FUNCTION_BLOCK FB_CIP_Client EXTENDS FB_SFC_Cycle IMPLEMENTS ITF_FB_SFC_Cycle
VAR_INPUT
	//eElementID			: E_Element_List;
	
	valClient_Source		: E_Pis_Name;
	valClient_Return		: E_Pis_Name;
	valS_Marinade_Up		: E_Pis_Name;
	//valS_Marinade_Up_Drain	: E_Pis_Name;
	valS_Marinade_Low		: E_Pis_Name;
	valS_Color_Up			: E_Pis_Name;
	//valS_Color_Up_Drain		: E_Pis_Name;
	valS_Color_Low			: E_Pis_Name;
	//valTank_1				: E_Pis_Name;
	//valTank_2				: E_Pis_Name;
	//valTank_3				: E_Pis_Name;
	//valTank_4				: E_Pis_Name;
	//valS_Marinade_Low_Select	: E_Pis_Name;
	//valS_Color_Low_Select	: E_Pis_Name;
	valDrain				: E_Pis_Name;
	valLoop					: E_Pis_Name;//V1030
	valS_Future				: E_Pis_Name;
	
END_VAR
VAR_OUTPUT
END_VAR
VAR
	//refElement		: REFERENCE TO FB_Element;
	//refState_Long		: REFERENCE TO E_Element_State_Long;
	eReq				: E_CIP_Client_Selector;
	eProcess			: E_CIP_Client_Selector;
	eStatus				: E_CIP_Client_Selector;
	
	fbPis					: FB_Piston;
	stPis_Client_Source			: REFERENCE TO ST_Piston;
	stPis_Client_Return			: REFERENCE TO ST_Piston;
	stPis_S_Marinade_Up			: REFERENCE TO ST_Piston;
	//stPis_S_Marinade_Up_Drain	: REFERENCE TO ST_Piston;
	stPis_S_Marinade_Low		: REFERENCE TO ST_Piston;
	stPis_S_Color_Up			: REFERENCE TO ST_Piston;
	//stPis_S_Color_Up_Drain		: REFERENCE TO ST_Piston;
	stPis_S_Color_Low			: REFERENCE TO ST_Piston;
	//stPis_Tank_1				: REFERENCE TO ST_Piston;
	//stPis_Tank_2				: REFERENCE TO ST_Piston;
	//stPis_Tank_3				: REFERENCE TO ST_Piston;
	//stPis_Tank_4				: REFERENCE TO ST_Piston;
	//stPis_S_Marinade_Low_Select	: REFERENCE TO ST_Piston;
	//stPis_S_Color_Low_Select	: REFERENCE TO ST_Piston;
	stPis_Drain					: REFERENCE TO ST_Piston;	
	stPis_Loop					: REFERENCE TO ST_Piston;//V1030
	stPis_S_Future				: REFERENCE TO ST_Piston;

	tonDrainTime: TON;
	
	rt_Req_Reset: R_TRIG;

END_VAR
VAR_IN_OUT


END_VAR

act_GetReference();

act_Oper();
IF NOT Init.x THEN;
	act_Status();
END_IF

tonDrainTime(PT:=T#1M, IN:=eStatus=E_CIP_Client_Selector.eDrain);
IF tonDrainTime.Q 
AND eReq=E_CIP_Client_Selector.eNone
AND eProcess=E_CIP_Client_Selector.eNone
THEN;
	eReq:=E_CIP_Client_Selector.eClose;
END_IF

m_Request_Reset(memo:=rt_Req_Reset);//rt_Req_Reset: R_TRIG;

ACTION _aClose_active:
bStepDone:=FALSE;
IF TRUE 
AND eStatus=E_CIP_Client_Selector.eClose
THEN;
	bStepDone:=TRUE;
END_IF
END_ACTION

ACTION _aClose_entry:
fbPis.m_SetByRecipe(stPis:=stPis_Client_Source, 		req:=E_Piston_Recipe_State.Release);
fbPis.m_SetByRecipe(stPis:=stPis_Client_Return, 		req:=E_Piston_Recipe_State.Release);
fbPis.m_SetByRecipe(stPis:=stPis_S_Marinade_Up, 		req:=E_Piston_Recipe_State.Release);
fbPis.m_SetByRecipe(stPis:=stPis_S_Marinade_Low, 		req:=E_Piston_Recipe_State.Release);
fbPis.m_SetByRecipe(stPis:=stPis_S_Color_Up, 			req:=E_Piston_Recipe_State.Release);
fbPis.m_SetByRecipe(stPis:=stPis_S_Color_Low, 			req:=E_Piston_Recipe_State.Release);
fbPis.m_SetByRecipe(stPis:=stPis_Drain, 				req:=E_Piston_Recipe_State.Release);
fbPis.m_SetByRecipe(stPis:=stPis_Loop, 					req:=E_Piston_Recipe_State.Release);
fbPis.m_SetByRecipe(stPis:=stPis_S_Future, 				req:=E_Piston_Recipe_State.Release);
END_ACTION

ACTION _aColor_Low_active:
bStepDone:=FALSE;
IF TRUE 
AND eStatus=E_CIP_Client_Selector.eColor_Low
THEN;
	bStepDone:=TRUE;
END_IF
END_ACTION

ACTION _aColor_Low_entry:
fbPis.m_SetByRecipe(stPis:=stPis_Client_Source, 		req:=E_Piston_Recipe_State.Act);
fbPis.m_SetByRecipe(stPis:=stPis_Client_Return, 		req:=E_Piston_Recipe_State.Act);
fbPis.m_SetByRecipe(stPis:=stPis_S_Marinade_Up, 		req:=E_Piston_Recipe_State.Release);
fbPis.m_SetByRecipe(stPis:=stPis_S_Marinade_Low, 		req:=E_Piston_Recipe_State.Release);
fbPis.m_SetByRecipe(stPis:=stPis_S_Color_Up, 			req:=E_Piston_Recipe_State.Release);
fbPis.m_SetByRecipe(stPis:=stPis_S_Color_Low, 			req:=E_Piston_Recipe_State.Act);
fbPis.m_SetByRecipe(stPis:=stPis_Drain, 				req:=E_Piston_Recipe_State.Release);
fbPis.m_SetByRecipe(stPis:=stPis_Loop, 					req:=E_Piston_Recipe_State.Release);
fbPis.m_SetByRecipe(stPis:=stPis_S_Future, 				req:=E_Piston_Recipe_State.Release);
END_ACTION

ACTION _aColor_Up_active:
bStepDone:=FALSE;
IF TRUE 
AND eStatus=E_CIP_Client_Selector.eColor_Up
THEN;
	bStepDone:=TRUE;
END_IF
END_ACTION

ACTION _aColor_Up_entry:
fbPis.m_SetByRecipe(stPis:=stPis_Client_Source, 		req:=E_Piston_Recipe_State.Act);
fbPis.m_SetByRecipe(stPis:=stPis_Client_Return, 		req:=E_Piston_Recipe_State.Act);
fbPis.m_SetByRecipe(stPis:=stPis_S_Marinade_Up, 		req:=E_Piston_Recipe_State.Release);
fbPis.m_SetByRecipe(stPis:=stPis_S_Marinade_Low, 		req:=E_Piston_Recipe_State.Release);
fbPis.m_SetByRecipe(stPis:=stPis_S_Color_Up, 			req:=E_Piston_Recipe_State.Act);
fbPis.m_SetByRecipe(stPis:=stPis_S_Color_Low, 			req:=E_Piston_Recipe_State.Release);
fbPis.m_SetByRecipe(stPis:=stPis_Drain, 				req:=E_Piston_Recipe_State.Release);
fbPis.m_SetByRecipe(stPis:=stPis_Loop, 					req:=E_Piston_Recipe_State.Release);
fbPis.m_SetByRecipe(stPis:=stPis_S_Future, 				req:=E_Piston_Recipe_State.Release);
END_ACTION

ACTION _aDone_entry:
eProcess:=E_CIP_Usage.eNotInUse;
eReq:=E_CIP_Usage.eNotInUse;
bRun:=FALSE;
bDone:=TRUE;
END_ACTION

ACTION _aDrain_active:
bStepDone:=FALSE;
IF TRUE 
AND eStatus=E_CIP_Client_Selector.eDrain
THEN;
	bStepDone:=TRUE;
END_IF
END_ACTION

ACTION _aDrain_entry:
fbPis.m_SetByRecipe(stPis:=stPis_Client_Source, 		req:=E_Piston_Recipe_State.Release);
fbPis.m_SetByRecipe(stPis:=stPis_Client_Return, 		req:=E_Piston_Recipe_State.Release);
fbPis.m_SetByRecipe(stPis:=stPis_S_Marinade_Up, 		req:=E_Piston_Recipe_State.Release);
fbPis.m_SetByRecipe(stPis:=stPis_S_Marinade_Low, 		req:=E_Piston_Recipe_State.Release);
fbPis.m_SetByRecipe(stPis:=stPis_S_Color_Up, 			req:=E_Piston_Recipe_State.Release);
fbPis.m_SetByRecipe(stPis:=stPis_S_Color_Low, 			req:=E_Piston_Recipe_State.Release);
fbPis.m_SetByRecipe(stPis:=stPis_Drain, 				req:=E_Piston_Recipe_State.Act);
fbPis.m_SetByRecipe(stPis:=stPis_Loop, 					req:=E_Piston_Recipe_State.Release);
fbPis.m_SetByRecipe(stPis:=stPis_S_Future, 				req:=E_Piston_Recipe_State.Release);
END_ACTION

ACTION _aFuture_active:
bStepDone:=FALSE;
IF TRUE 
AND eStatus=E_CIP_Client_Selector.eFuture
THEN;
	bStepDone:=TRUE;
END_IF
END_ACTION

ACTION _aFuture_entry:
fbPis.m_SetByRecipe(stPis:=stPis_Client_Source, 		req:=E_Piston_Recipe_State.Act);
fbPis.m_SetByRecipe(stPis:=stPis_Client_Return, 		req:=E_Piston_Recipe_State.Act);
fbPis.m_SetByRecipe(stPis:=stPis_S_Marinade_Up, 		req:=E_Piston_Recipe_State.Release);
fbPis.m_SetByRecipe(stPis:=stPis_S_Marinade_Low, 		req:=E_Piston_Recipe_State.Release);
fbPis.m_SetByRecipe(stPis:=stPis_S_Color_Up, 			req:=E_Piston_Recipe_State.Release);
fbPis.m_SetByRecipe(stPis:=stPis_S_Color_Low, 			req:=E_Piston_Recipe_State.Release);
fbPis.m_SetByRecipe(stPis:=stPis_Drain, 				req:=E_Piston_Recipe_State.Release);
fbPis.m_SetByRecipe(stPis:=stPis_Loop, 					req:=E_Piston_Recipe_State.Release);
fbPis.m_SetByRecipe(stPis:=stPis_S_Future, 				req:=E_Piston_Recipe_State.Act);
END_ACTION

ACTION _aInit_active:
SFCReset:=FALSE;
END_ACTION

ACTION _aInit_exit:
eProcess:=E_CIP_Usage.eNotInUse;
eReq:=E_CIP_Usage.eNotInUse;
END_ACTION

ACTION _aLoop_active:
bStepDone:=FALSE;
IF TRUE 
AND eStatus=E_CIP_Client_Selector.eLoop
THEN;
	bStepDone:=TRUE;
END_IF
END_ACTION

ACTION _aLoop_entry:
fbPis.m_SetByRecipe(stPis:=stPis_Client_Source, 		req:=E_Piston_Recipe_State.Act);
fbPis.m_SetByRecipe(stPis:=stPis_Client_Return, 		req:=E_Piston_Recipe_State.Act);
fbPis.m_SetByRecipe(stPis:=stPis_S_Marinade_Up, 		req:=E_Piston_Recipe_State.Release);
fbPis.m_SetByRecipe(stPis:=stPis_S_Marinade_Low, 		req:=E_Piston_Recipe_State.Release);
fbPis.m_SetByRecipe(stPis:=stPis_S_Color_Up, 			req:=E_Piston_Recipe_State.Release);
fbPis.m_SetByRecipe(stPis:=stPis_S_Color_Low, 			req:=E_Piston_Recipe_State.Release);
fbPis.m_SetByRecipe(stPis:=stPis_Drain, 				req:=E_Piston_Recipe_State.Act);
fbPis.m_SetByRecipe(stPis:=stPis_Loop, 					req:=E_Piston_Recipe_State.Act);
fbPis.m_SetByRecipe(stPis:=stPis_S_Future, 				req:=E_Piston_Recipe_State.Release);
END_ACTION

ACTION _aMarinade_Low_active:
bStepDone:=FALSE;
IF TRUE 
AND eStatus=E_CIP_Client_Selector.eMarinade_Low
THEN;
	bStepDone:=TRUE;
END_IF
END_ACTION

ACTION _aMarinade_Low_entry:
fbPis.m_SetByRecipe(stPis:=stPis_Client_Source, 		req:=E_Piston_Recipe_State.Act);
fbPis.m_SetByRecipe(stPis:=stPis_Client_Return, 		req:=E_Piston_Recipe_State.Act);
fbPis.m_SetByRecipe(stPis:=stPis_S_Marinade_Up, 		req:=E_Piston_Recipe_State.Release);
fbPis.m_SetByRecipe(stPis:=stPis_S_Marinade_Low, 		req:=E_Piston_Recipe_State.Act);
fbPis.m_SetByRecipe(stPis:=stPis_S_Color_Up, 			req:=E_Piston_Recipe_State.Release);
fbPis.m_SetByRecipe(stPis:=stPis_S_Color_Low, 			req:=E_Piston_Recipe_State.Release);
fbPis.m_SetByRecipe(stPis:=stPis_Drain, 				req:=E_Piston_Recipe_State.Release);
fbPis.m_SetByRecipe(stPis:=stPis_Loop, 					req:=E_Piston_Recipe_State.Release);
fbPis.m_SetByRecipe(stPis:=stPis_S_Future, 				req:=E_Piston_Recipe_State.Release);
END_ACTION

ACTION _aMarinade_Up_active:
bStepDone:=FALSE;
IF TRUE 
AND eStatus=E_CIP_Client_Selector.eMarinade_Up
THEN;
	bStepDone:=TRUE;
END_IF
END_ACTION

ACTION _aMarinade_Up_entry:
fbPis.m_SetByRecipe(stPis:=stPis_Client_Source, 		req:=E_Piston_Recipe_State.Act);
fbPis.m_SetByRecipe(stPis:=stPis_Client_Return, 		req:=E_Piston_Recipe_State.Act);
fbPis.m_SetByRecipe(stPis:=stPis_S_Marinade_Up, 		req:=E_Piston_Recipe_State.Act);
fbPis.m_SetByRecipe(stPis:=stPis_S_Marinade_Low, 		req:=E_Piston_Recipe_State.Release);
fbPis.m_SetByRecipe(stPis:=stPis_S_Color_Up, 			req:=E_Piston_Recipe_State.Release);
fbPis.m_SetByRecipe(stPis:=stPis_S_Color_Low, 			req:=E_Piston_Recipe_State.Release);
fbPis.m_SetByRecipe(stPis:=stPis_Drain, 				req:=E_Piston_Recipe_State.Release);
fbPis.m_SetByRecipe(stPis:=stPis_Loop, 					req:=E_Piston_Recipe_State.Release);
fbPis.m_SetByRecipe(stPis:=stPis_S_Future, 				req:=E_Piston_Recipe_State.Release);
END_ACTION

ACTION _aReady_active:


IF eReq<>E_CIP_Client_Selector.eNone THEN;
	IF eProcess=E_CIP_Client_Selector.eNone 
	THEN;
		eProcess:=eReq;
	ELSE;
		eReq:=E_CIP_Client_Selector.eNone;
	END_IF
END_IF

(*
CASE eReq OF
	E_CIP_Usage.eLine_Color:;
			IF TRUE THEN;
				eProcess:=E_CIP_Usage.eLine_Color;
			END_IF

	E_CIP_Usage.eLine_Marinada:;
			IF TRUE THEN;
				eProcess:=E_CIP_Usage.eLine_Marinada;
			END_IF	
			
	E_CIP_Usage.eLocal:;
			IF TRUE THEN;
				eProcess:=E_CIP_Usage.eLocal;
			END_IF	

	E_CIP_Usage.eNotInUse:;
			IF TRUE THEN;
				eProcess:=E_CIP_Usage.eNotInUse;
			END_IF	
			
	E_CIP_Usage.eTank_1:;
			IF TRUE THEN;
				eProcess:=E_CIP_Usage.eTank_1;
			END_IF	
	E_CIP_Usage.eTank_2:;
			IF TRUE THEN;
				eProcess:=E_CIP_Usage.eTank_2;
			END_IF	
	E_CIP_Usage.eTank_3:;
			IF TRUE THEN;
				eProcess:=E_CIP_Usage.eTank_3;
			END_IF	
	E_CIP_Usage.eTank_4:;
			IF TRUE THEN;
				eProcess:=E_CIP_Usage.eTank_4;
			END_IF	
	E_CIP_Usage.eTriBlender_Color:;
			IF TRUE THEN;
				eProcess:=E_CIP_Usage.eTriBlender_Color;
			END_IF	
	E_CIP_Usage.eTriBlender_Marinada:;
			IF TRUE THEN;
				eProcess:=E_CIP_Usage.eTriBlender_Marinada;
			END_IF	

END_CASE
*)
END_ACTION

ACTION _aReady_exit:
bRun:=TRUE;
bDone:=FALSE;
END_ACTION

ACTION act_GetReference:
m_Set_SFCFlags_Reference();
//refElement REF= fbElement[eElementID];
//refState_Long REF= fbElement[eElementID].eState_Long;

stPis_Client_Source			REF= g_Piston.stPis[valClient_Source];
stPis_Client_Return			REF= g_Piston.stPis[valClient_Return];
stPis_S_Marinade_Up			REF= g_Piston.stPis[valS_Marinade_Up];
//stPis_S_Marinade_Up_Drain	REF= g_Piston.stPis[valS_Marinade_Up_Drain];
stPis_S_Marinade_Low		REF= g_Piston.stPis[valS_Marinade_Low];
stPis_S_Color_Up			REF= g_Piston.stPis[valS_Color_Up];
//stPis_S_Color_Up_Drain		REF= g_Piston.stPis[valS_Color_Up_Drain];
stPis_S_Color_Low			REF= g_Piston.stPis[valS_Color_Low];
//stPis_Tank_1				REF= g_Piston.stPis[valTank_1];
//stPis_Tank_2				REF= g_Piston.stPis[valTank_2];
//stPis_Tank_3				REF= g_Piston.stPis[valTank_3];
//stPis_Tank_4				REF= g_Piston.stPis[valTank_4];
//stPis_S_Marinade_Low_Select	REF= g_Piston.stPis[valS_Marinade_Low_Select];
//stPis_S_Color_Low_Select	REF= g_Piston.stPis[valS_Color_Low_Select];
stPis_Drain					REF= g_Piston.stPis[valDrain];
stPis_Loop				REF= g_Piston.stPis[valLoop];
stPis_S_Future				REF= g_Piston.stPis[valS_Future];
END_ACTION

ACTION act_Oper:
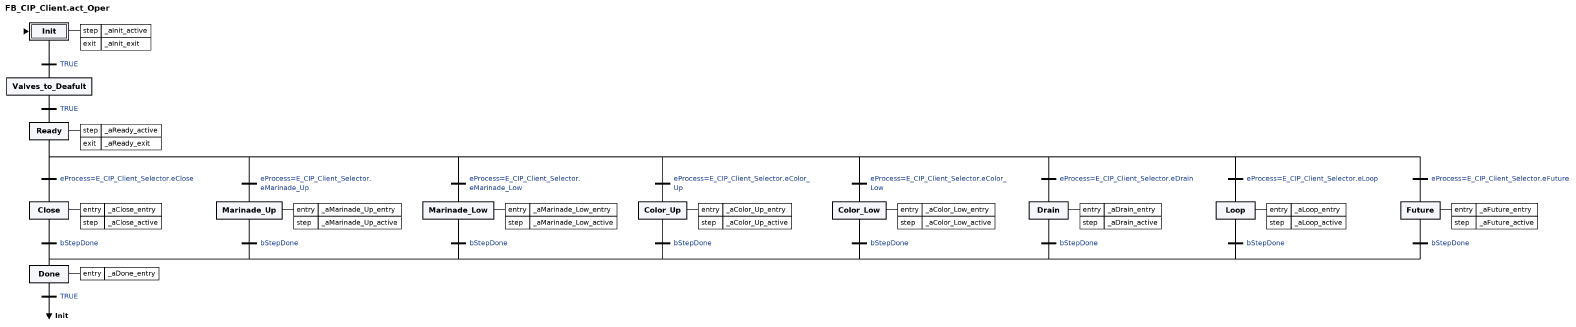
INITIAL_STEP Init:  // min time T#0.5s
    _aInit_active(N);  // step action
    _aInit_exit(P0);  // exit action
END_STEP
TRANSITION FROM Init TO Valves_to_Deafult
    := TRUE;
END_TRANSITION
STEP Valves_to_Deafult:
END_STEP
TRANSITION FROM Valves_to_Deafult TO Ready
    := TRUE;
END_TRANSITION
STEP Ready:
    _aReady_active(N);  // step action
    _aReady_exit(P0);  // exit action
END_STEP
TRANSITION FROM Ready TO Close
    := eProcess=E_CIP_Client_Selector.eClose;
END_TRANSITION
STEP Close:
    _aClose_entry(P1);  // entry action
    _aClose_active(N);  // step action
END_STEP
TRANSITION FROM Close TO Done
    := bStepDone;
END_TRANSITION
TRANSITION FROM Ready TO Marinade_Up
    := eProcess=E_CIP_Client_Selector.eMarinade_Up;
END_TRANSITION
STEP Marinade_Up:
    _aMarinade_Up_entry(P1);  // entry action
    _aMarinade_Up_active(N);  // step action
END_STEP
TRANSITION FROM Marinade_Up TO Done
    := bStepDone;
END_TRANSITION
TRANSITION FROM Ready TO Marinade_Low
    := eProcess=E_CIP_Client_Selector.eMarinade_Low;
END_TRANSITION
STEP Marinade_Low:
    _aMarinade_Low_entry(P1);  // entry action
    _aMarinade_Low_active(N);  // step action
END_STEP
TRANSITION FROM Marinade_Low TO Done
    := bStepDone;
END_TRANSITION
TRANSITION FROM Ready TO Color_Up
    := eProcess=E_CIP_Client_Selector.eColor_Up;
END_TRANSITION
STEP Color_Up:
    _aColor_Up_entry(P1);  // entry action
    _aColor_Up_active(N);  // step action
END_STEP
TRANSITION FROM Color_Up TO Done
    := bStepDone;
END_TRANSITION
TRANSITION FROM Ready TO Color_Low
    := eProcess=E_CIP_Client_Selector.eColor_Low;
END_TRANSITION
STEP Color_Low:
    _aColor_Low_entry(P1);  // entry action
    _aColor_Low_active(N);  // step action
END_STEP
TRANSITION FROM Color_Low TO Done
    := bStepDone;
END_TRANSITION
TRANSITION FROM Ready TO Drain
    := eProcess=E_CIP_Client_Selector.eDrain;
END_TRANSITION
STEP Drain:
    _aDrain_entry(P1);  // entry action
    _aDrain_active(N);  // step action
END_STEP
TRANSITION FROM Drain TO Done
    := bStepDone;
END_TRANSITION
TRANSITION FROM Ready TO Loop
    := eProcess=E_CIP_Client_Selector.eLoop;
END_TRANSITION
STEP Loop:
    _aLoop_entry(P1);  // entry action
    _aLoop_active(N);  // step action
END_STEP
TRANSITION FROM Loop TO Done
    := bStepDone;
END_TRANSITION
TRANSITION FROM Ready TO Future
    := eProcess=E_CIP_Client_Selector.eFuture;
END_TRANSITION
STEP Future:
    _aFuture_entry(P1);  // entry action
    _aFuture_active(N);  // step action
END_STEP
TRANSITION FROM Future TO Done
    := bStepDone;
END_TRANSITION
STEP Done:  // min time T#0.2s
    _aDone_entry(P1);  // entry action
END_STEP
TRANSITION FROM Done TO Init
    := TRUE;
END_TRANSITION
// branch label Branch2_act_Oper
END_ACTION

ACTION act_Status:
IF bReady AND bDone OR TRUE THEN;
	IF TRUE 
	AND fbPis.m_CheckByRecipe(stPis:=stPis_Client_Source, 		req:=E_Piston_Recipe_State.Release)
	AND fbPis.m_CheckByRecipe(stPis:=stPis_Client_Return, 		req:=E_Piston_Recipe_State.Release)
	AND fbPis.m_CheckByRecipe(stPis:=stPis_S_Marinade_Up, 		req:=E_Piston_Recipe_State.Release)
	AND fbPis.m_CheckByRecipe(stPis:=stPis_S_Marinade_Low, 		req:=E_Piston_Recipe_State.Release)
	AND fbPis.m_CheckByRecipe(stPis:=stPis_S_Color_Up, 			req:=E_Piston_Recipe_State.Release)
	AND fbPis.m_CheckByRecipe(stPis:=stPis_S_Color_Low, 		req:=E_Piston_Recipe_State.Release)
	AND fbPis.m_CheckByRecipe(stPis:=stPis_Drain, 				req:=E_Piston_Recipe_State.Release)
	AND fbPis.m_CheckByRecipe(stPis:=stPis_Loop, 				req:=E_Piston_Recipe_State.Release)
	AND fbPis.m_CheckByRecipe(stPis:=stPis_S_Future, 			req:=E_Piston_Recipe_State.Release)
	THEN;
		eStatus:=E_CIP_Client_Selector.eClose;
	ELSIF TRUE
	AND fbPis.m_CheckByRecipe(stPis:=stPis_Client_Source, 		req:=E_Piston_Recipe_State.Act)
	AND fbPis.m_CheckByRecipe(stPis:=stPis_Client_Return, 		req:=E_Piston_Recipe_State.Act)
	AND fbPis.m_CheckByRecipe(stPis:=stPis_S_Marinade_Up, 		req:=E_Piston_Recipe_State.Act)
	AND fbPis.m_CheckByRecipe(stPis:=stPis_S_Marinade_Low, 		req:=E_Piston_Recipe_State.Release)
	AND fbPis.m_CheckByRecipe(stPis:=stPis_S_Color_Up, 			req:=E_Piston_Recipe_State.Release)
	AND fbPis.m_CheckByRecipe(stPis:=stPis_S_Color_Low, 		req:=E_Piston_Recipe_State.Release)
	AND fbPis.m_CheckByRecipe(stPis:=stPis_Drain, 				req:=E_Piston_Recipe_State.Release)
	AND fbPis.m_CheckByRecipe(stPis:=stPis_Loop, 				req:=E_Piston_Recipe_State.Release)
	AND fbPis.m_CheckByRecipe(stPis:=stPis_S_Future, 			req:=E_Piston_Recipe_State.Release)
	THEN;
		eStatus:=E_CIP_Client_Selector.eMarinade_Up;
	ELSIF TRUE 
	AND fbPis.m_CheckByRecipe(stPis:=stPis_Client_Source, 		req:=E_Piston_Recipe_State.Act)
	AND fbPis.m_CheckByRecipe(stPis:=stPis_Client_Return, 		req:=E_Piston_Recipe_State.Act)
	AND fbPis.m_CheckByRecipe(stPis:=stPis_S_Marinade_Up, 		req:=E_Piston_Recipe_State.Release)
	AND fbPis.m_CheckByRecipe(stPis:=stPis_S_Marinade_Low, 		req:=E_Piston_Recipe_State.Act)
	AND fbPis.m_CheckByRecipe(stPis:=stPis_S_Color_Up, 			req:=E_Piston_Recipe_State.Release)
	AND fbPis.m_CheckByRecipe(stPis:=stPis_S_Color_Low, 		req:=E_Piston_Recipe_State.Release)
	AND fbPis.m_CheckByRecipe(stPis:=stPis_Drain, 				req:=E_Piston_Recipe_State.Release)
	AND fbPis.m_CheckByRecipe(stPis:=stPis_Loop, 				req:=E_Piston_Recipe_State.Release)
	AND fbPis.m_CheckByRecipe(stPis:=stPis_S_Future, 			req:=E_Piston_Recipe_State.Release)
	THEN;
		eStatus:=E_CIP_Client_Selector.eMarinade_Low;
	ELSIF TRUE 
	AND fbPis.m_CheckByRecipe(stPis:=stPis_Client_Source, 		req:=E_Piston_Recipe_State.Act)
	AND fbPis.m_CheckByRecipe(stPis:=stPis_Client_Return, 		req:=E_Piston_Recipe_State.Act)
	AND fbPis.m_CheckByRecipe(stPis:=stPis_S_Marinade_Up, 		req:=E_Piston_Recipe_State.Release)
	AND fbPis.m_CheckByRecipe(stPis:=stPis_S_Marinade_Low, 		req:=E_Piston_Recipe_State.Release)
	AND fbPis.m_CheckByRecipe(stPis:=stPis_S_Color_Up, 			req:=E_Piston_Recipe_State.Act)
	AND fbPis.m_CheckByRecipe(stPis:=stPis_S_Color_Low, 		req:=E_Piston_Recipe_State.Release)
	AND fbPis.m_CheckByRecipe(stPis:=stPis_Drain, 				req:=E_Piston_Recipe_State.Release)
	AND fbPis.m_CheckByRecipe(stPis:=stPis_Loop, 				req:=E_Piston_Recipe_State.Release)
	AND fbPis.m_CheckByRecipe(stPis:=stPis_S_Future, 			req:=E_Piston_Recipe_State.Release)
	THEN;
		eStatus:=E_CIP_Client_Selector.eColor_Up;
	ELSIF TRUE 
	AND fbPis.m_CheckByRecipe(stPis:=stPis_Client_Source, 		req:=E_Piston_Recipe_State.Act)
	AND fbPis.m_CheckByRecipe(stPis:=stPis_Client_Return, 		req:=E_Piston_Recipe_State.Act)
	AND fbPis.m_CheckByRecipe(stPis:=stPis_S_Marinade_Up, 		req:=E_Piston_Recipe_State.Release)
	AND fbPis.m_CheckByRecipe(stPis:=stPis_S_Marinade_Low, 		req:=E_Piston_Recipe_State.Release)
	AND fbPis.m_CheckByRecipe(stPis:=stPis_S_Color_Up, 			req:=E_Piston_Recipe_State.Release)
	AND fbPis.m_CheckByRecipe(stPis:=stPis_S_Color_Low, 		req:=E_Piston_Recipe_State.Act)
	AND fbPis.m_CheckByRecipe(stPis:=stPis_Drain, 				req:=E_Piston_Recipe_State.Release)
	AND fbPis.m_CheckByRecipe(stPis:=stPis_Loop, 				req:=E_Piston_Recipe_State.Release)
	AND fbPis.m_CheckByRecipe(stPis:=stPis_S_Future, 			req:=E_Piston_Recipe_State.Release)
	THEN;
		eStatus:=E_CIP_Client_Selector.eColor_Low;
	ELSIF TRUE 
	AND fbPis.m_CheckByRecipe(stPis:=stPis_Client_Source, 		req:=E_Piston_Recipe_State.Release)
	AND fbPis.m_CheckByRecipe(stPis:=stPis_Client_Return, 		req:=E_Piston_Recipe_State.Release)
	AND fbPis.m_CheckByRecipe(stPis:=stPis_S_Marinade_Up, 		req:=E_Piston_Recipe_State.Release)
	AND fbPis.m_CheckByRecipe(stPis:=stPis_S_Marinade_Low, 		req:=E_Piston_Recipe_State.Release)
	AND fbPis.m_CheckByRecipe(stPis:=stPis_S_Color_Up, 			req:=E_Piston_Recipe_State.Release)
	AND fbPis.m_CheckByRecipe(stPis:=stPis_S_Color_Low, 		req:=E_Piston_Recipe_State.Release)
	AND fbPis.m_CheckByRecipe(stPis:=stPis_Drain, 				req:=E_Piston_Recipe_State.Act)
	AND fbPis.m_CheckByRecipe(stPis:=stPis_Loop, 				req:=E_Piston_Recipe_State.Release)
	AND fbPis.m_CheckByRecipe(stPis:=stPis_S_Future, 			req:=E_Piston_Recipe_State.Release)
	THEN;
		eStatus:=E_CIP_Client_Selector.eDrain;
	ELSIF TRUE 
	AND fbPis.m_CheckByRecipe(stPis:=stPis_Client_Source, 		req:=E_Piston_Recipe_State.Act)
	AND fbPis.m_CheckByRecipe(stPis:=stPis_Client_Return, 		req:=E_Piston_Recipe_State.Act)
	AND fbPis.m_CheckByRecipe(stPis:=stPis_S_Marinade_Up, 		req:=E_Piston_Recipe_State.Release)
	AND fbPis.m_CheckByRecipe(stPis:=stPis_S_Marinade_Low, 		req:=E_Piston_Recipe_State.Release)
	AND fbPis.m_CheckByRecipe(stPis:=stPis_S_Color_Up, 			req:=E_Piston_Recipe_State.Release)
	AND fbPis.m_CheckByRecipe(stPis:=stPis_S_Color_Low, 		req:=E_Piston_Recipe_State.Release)
	AND fbPis.m_CheckByRecipe(stPis:=stPis_Drain, 				req:=E_Piston_Recipe_State.Act)
	AND fbPis.m_CheckByRecipe(stPis:=stPis_Loop, 				req:=E_Piston_Recipe_State.Act)
	AND fbPis.m_CheckByRecipe(stPis:=stPis_S_Future, 			req:=E_Piston_Recipe_State.Release)
	THEN;
		eStatus:=E_CIP_Client_Selector.eLoop;
	ELSIF TRUE 
	AND fbPis.m_CheckByRecipe(stPis:=stPis_Client_Source, 		req:=E_Piston_Recipe_State.Act)
	AND fbPis.m_CheckByRecipe(stPis:=stPis_Client_Return, 		req:=E_Piston_Recipe_State.Act)
	AND fbPis.m_CheckByRecipe(stPis:=stPis_S_Marinade_Up, 		req:=E_Piston_Recipe_State.Release)
	AND fbPis.m_CheckByRecipe(stPis:=stPis_S_Marinade_Low, 		req:=E_Piston_Recipe_State.Release)
	AND fbPis.m_CheckByRecipe(stPis:=stPis_S_Color_Up, 			req:=E_Piston_Recipe_State.Release)
	AND fbPis.m_CheckByRecipe(stPis:=stPis_S_Color_Low, 		req:=E_Piston_Recipe_State.Release)
	AND fbPis.m_CheckByRecipe(stPis:=stPis_Drain, 				req:=E_Piston_Recipe_State.Release)
	AND fbPis.m_CheckByRecipe(stPis:=stPis_Loop, 				req:=E_Piston_Recipe_State.Release)
	AND fbPis.m_CheckByRecipe(stPis:=stPis_S_Future, 			req:=E_Piston_Recipe_State.Act)
	THEN;
		eStatus:=E_CIP_Client_Selector.eFuture;
	ELSE;
		eStatus:=E_CIP_Client_Selector.eNone;
	END_IF
ELSE;
	eStatus:=E_CIP_Client_Selector.eNone;
END_IF
END_ACTION

METHOD m_CheckStatus : BOOL
VAR_INPUT
	eReqStatus		: E_CIP_Usage;
END_VAR
VAR
	eReqStatusLocal	: E_CIP_Client_Selector;
END_VAR
CASE eReqStatus OF
	E_CIP_Usage.eLocal:;
				eReqStatusLocal	:=E_CIP_Client_Selector.eClose;
	E_CIP_Usage.eTank_1,
	E_CIP_Usage.eTank_2:;
				eReqStatusLocal	:=E_CIP_Client_Selector.eMarinade_Up;	
	E_CIP_Usage.eTank_3,
	E_CIP_Usage.eTank_4:;
				eReqStatusLocal	:=E_CIP_Client_Selector.eColor_Up;	
	E_CIP_Usage.eTriBlender_Marinada,
	E_CIP_Usage.eLine_Marinada:;
				eReqStatusLocal	:=E_CIP_Client_Selector.eMarinade_Low;	
	E_CIP_Usage.eTriBlender_Color,
	E_CIP_Usage.eLine_Color:;
				eReqStatusLocal	:=E_CIP_Client_Selector.eColor_Low;	
	
END_CASE

IF eStatus=eReqStatusLocal 
AND eProcess=E_CIP_Client_Selector.eNone
AND eReq=E_CIP_Client_Selector.eNone
AND bReady
AND bDone
AND NOT bRun
THEN;
	m_CheckStatus:=TRUE;
END_IF
END_METHOD

METHOD m_Request_Reset : BOOL
VAR_IN_OUT
	memo: R_TRIG;
END_VAR
memo(CLK:=eReq=0);
IF TRUE 
AND memo.Q
THEN;
	SFCReset:=TRUE;
END_IF
END_METHOD

METHOD m_Run : BOOL
VAR_INPUT
	eReqProc			: E_CIP_Usage;
END_VAR
VAR
	eReqStatusLocal	: E_CIP_Client_Selector;
END_VAR
CASE eReqProc OF
	E_CIP_Usage.eLocal:;
				eReqStatusLocal	:=E_CIP_Client_Selector.eClose;
	E_CIP_Usage.eTank_1,
	E_CIP_Usage.eTank_2:;
				eReqStatusLocal	:=E_CIP_Client_Selector.eMarinade_Up;	
	E_CIP_Usage.eTank_3,
	E_CIP_Usage.eTank_4:;
				eReqStatusLocal	:=E_CIP_Client_Selector.eColor_Up;	
	E_CIP_Usage.eTriBlender_Marinada,
	E_CIP_Usage.eLine_Marinada:;
				eReqStatusLocal	:=E_CIP_Client_Selector.eMarinade_Low;	
	E_CIP_Usage.eTriBlender_Color,
	E_CIP_Usage.eLine_Color:;
				eReqStatusLocal	:=E_CIP_Client_Selector.eColor_Low;	
	
END_CASE

IF eProcess=E_CIP_Client_Selector.eNone THEN;
	eProcess:=eReq:=eReqStatusLocal;
	bDone:=FALSE;
	m_Run:=TRUE;
END_IF
END_METHOD

METHOD m_Set_SFCFlags_Reference : BOOL
//Set reference to SFC flags

refSFC.SFCInit REF= SFCInit;
refSFC.SFCReset REF= SFCReset;
refSFC.SFCError REF= SFCError;
refSFC.SFCEnableLimit REF= SFCEnableLimit;
refSFC.SFCErrorStep REF= SFCErrorStep;
refSFC.SFCErrorPOU REF= SFCErrorPOU;
refSFC.SFCQuitError REF= SFCQuitError;
refSFC.SFCPause REF= SFCPause;
refSFC.SFCTrans REF= SFCTrans;
refSFC.SFCCurrentStep REF= SFCCurrentStep;
refSFC.SFCTip REF= SFCTip;
refSFC.SFCTipMode REF= SFCTipMode;

// Cycle handle for SFC
m_SFC_Handle();
END_METHOD

END_FUNCTION_BLOCK

(* stored: Version 1.1.0.1, ProductVersion 3.1.4024.13
   POU FB_CIP_Client: Id {c5033c12-cb76-4d9f-9912-a992211c6f9c}, SpecialFunc None
   Folder Manage: Id {38103117-043f-403d-a53b-cc92b5c9eca8}
   Action _aClose_active: Id {0c273ec4-07ea-4c3a-9a5b-c8ebfdd77695}
   Action _aClose_entry: Id {89bb949b-73b9-4e77-8017-b6327b0bdda0}
   Action _aColor_Low_active: Id {88414d37-f878-422b-978f-18c0dc12a666}
   Action _aColor_Low_entry: Id {c1927158-4d78-451e-a925-f4404ebed7c3}
   Action _aColor_Up_active: Id {371c6bec-9334-4491-864a-d33c65b63a61}
   Action _aColor_Up_entry: Id {28e65717-9ec3-49b4-9c7a-55f22afa9837}
   Action _aDone_entry: Id {60428b5e-2664-48fc-baa3-5f1fc5212655}
   Action _aDrain_active: Id {72cc4ab0-083a-4817-a202-7c56b859c63c}
   Action _aDrain_entry: Id {954a9e30-8407-40fd-8169-d919834d753b}
   Action _aFuture_active: Id {74285a53-17ed-49d1-8065-636d4e3f572f}
   Action _aFuture_entry: Id {8f148dfe-1383-4cb1-b559-71eda112affa}
   Action _aInit_active: Id {ba4548f9-0bde-4457-a942-f84ef37dcc1c}
   Action _aInit_exit: Id {f29be3ee-e528-4005-96b2-1ef3343e2f94}
   Action _aLoop_active: Id {3c0e8be8-f6f7-4fe6-b7ac-8c6a37c70621}
   Action _aLoop_entry: Id {c991bc47-9ace-4a84-884a-f03475ca6c26}
   Action _aMarinade_Low_active: Id {d1483e64-4746-49a3-9e31-99ca013c3759}
   Action _aMarinade_Low_entry: Id {14fd1617-abf4-47e8-b906-b9c9df5f476d}
   Action _aMarinade_Up_active: Id {35ac2ee3-7118-443b-9114-b224b600d3b5}
   Action _aMarinade_Up_entry: Id {328f52ec-1b83-47ac-84bf-d158e139b2f9}
   Action _aReady_active: Id {08fcf68e-dc0f-47ca-acbd-f456115322bd}
   Action _aReady_exit: Id {5f3f3241-71ef-4f6c-8d41-41776643de15}
   Action act_GetReference: Id {84cac95e-a105-49db-a8ae-c6f6784af55d}
   Action act_Oper: Id {ed4bd9f9-7bcc-429e-a8d9-d36dd2b5f0b3}
   Action act_Status: Id {62143100-fdee-42d6-8a63-1ad3f74db813}
   Method m_CheckStatus: Id {b5de556e-91b0-4df7-96d4-bc419ec06c1d}
   Method m_Request_Reset: Id {3a0085ac-d519-46ef-8977-d86d9a880e6b}
   Method m_Run: Id {a8bdb2df-eb11-4961-9b0c-b01d07d5677a}
   Method m_Set_SFCFlags_Reference: Id {6740c604-b51a-4401-88e7-e8f7ceec239c} *)
